(* IEC 61131-3 sources: codesys-framework/txt/application/ToDo/Hardware/IO/Cylinder/FB_Cylinder/Private, 5 files *)

(* ---- ProcessDetections.method.st ---- *)
METHOD PROTECTED ProcessDetections : BOOL
VAR_INPUT
END_VAR

// --- BEGIN IMPLEMENTATION ---

IF _eState = E_CylinderStates.GoToPos0
	AND ((_scSysPar.xSensorPresentPos0 AND _xDetPos0) OR (NOT _scSysPar.xSensorPresentPos0 AND _tonToPos0.Q))
THEN
	_eState := E_CylinderStates.Pos0;
END_IF

IF	_eState = E_CylinderStates.GoToPos1
	AND	((_scSysPar.xSensorPresentPos1 AND _xDetPos1) OR (NOT _scSysPar.xSensorPresentPos1 AND _tontopos1.Q))
THEN
	_eState := E_CylinderStates.Pos1;
END_IF

(* ---- ProcessErrors.method.st ---- *)
METHOD PROTECTED ProcessErrors
VAR_INPUT
END_VAR

// --- BEGIN IMPLEMENTATION ---

IF _scSysPar.xSensorPresentPos0 AND _tonToPos0.Q THEN

	_eState := E_CylinderStates.Invalid;
	_scError.xErrorActive := TRUE;
	_scError.sError := CONCAT(_sName, ': did not reach position 0 in time.');

END_IF

IF _scSysPar.xSensorPresentPos1 AND _tonToPos1.Q THEN

	_eState := E_CylinderStates.Invalid;
	_scError.xErrorActive := TRUE;
	_scError.sError := CONCAT(_sName, ': did not reach position 1 in time.');

END_IF

IF _eState <> E_CylinderStates.Invalid THEN
	_scError.xErrorActive := FALSE;
	_scError.sError := '';
END_IF

(* ---- ProcessGoToPos0.method.st ---- *)
METHOD PROTECTED ProcessGoToPos0 : BOOL
VAR_INPUT
END_VAR

// --- BEGIN IMPLEMENTATION ---

xDQ_Value := FALSE;

(* ---- ProcessGoToPos1.method.st ---- *)
METHOD PRIVATE ProcessGoToPos1 : BOOL
VAR_INPUT
END_VAR

// --- BEGIN IMPLEMENTATION ---

xDQ_Value := TRUE;

(* ---- ProcessState.method.st ---- *)
METHOD PROTECTED ProcessState : BOOL
VAR_INPUT
END_VAR

// --- BEGIN IMPLEMENTATION ---

CASE _eState OF

	E_CylinderStates.Invalid		: ;
	E_CylinderStates.Pos0			: ;
	E_CylinderStates.Pos1			: ;
	E_CylinderStates.GoToPos0		: ProcessGoToPos0();
	E_CylinderStates.GoToPos1		: ProcessGoToPos1();

END_CASE

_xDone := _eState = E_CylinderStates.Pos0 OR _eState = E_CylinderStates.Pos1;
_xBusy := _eState = E_CylinderStates.GoToPos0 OR _eState = E_CylinderStates.GoToPos1;
